FUNCTION_BLOCK TcoContextTest EXTENDS TcoCore._internals_TcoContext
VAR
	_callMyPlcInstance 		:	BOOL := FALSE;
	_startCycles			:	ULINT;
	_endCycles				:	ULINT;	
	_mainCycles				:	ULINT;
	_tcoObjectTest_A		:	TcoObjectTest(THIS^);
	_tcoObjectTest_B		:	TcoObjectTest(THIS^);
	_tcoObjectTest_Misc		:	TcoObjectTest(THIS^);
	_myIdentity				:	ULINT;	
	_onEntryCount			:	ULINT;
	_onExitCount			:	ULINT;
END_VAR

IF THIS^._callMyPlcInstance THEN
	THIS^.Run();
END_IF

{attribute 'TcRpcEnable'}
METHOD INTERNAL CallMainFromUnitTest
THIS^.Main();
END_METHOD

{attribute 'TcRpcEnable'}
METHOD INTERNAL CallRunFromUnitTest
THIS^.Run();
END_METHOD

{attribute 'TcRpcEnable'}
METHOD INTERNAL ContextClose
SUPER^._Close();
END_METHOD

{attribute 'TcRpcEnable'}
METHOD INTERNAL ContextOpen
SUPER^._Open();
END_METHOD

METHOD PROTECTED  Main
_mainCycles := _mainCycles + 1;

_myIdentity	:= THIS^.Identity;
END_METHOD

(*~
	<docu>
		<summary>
			Called on entry into context. When overridden in derived class allows to execute an arbitrary logic prior to opening the context cycle.
			<remarks>			
				<note type="important">					
					The method executes prior to opening the context. The context might not be properly initialized on first call. 
					Any information contained in the context at this point are from the last execution.
				</note>
			</remarks>
		</summary>			
	</docu>	
~*)
METHOD PROTECTED OnEntry
_onEntryCount := _onEntryCount + 1;
END_METHOD


(*~
	<docu>
		<summary>
			Called upon exit from the context. When overridden in derived class allows to execute an arbitrary logic after closing the context cycle.	
		</summary>			
	</docu>	
~*)METHOD PROTECTED OnExit
_onExitCount := _onExitCount + 1;
END_METHOD

{attribute 'TcRpcEnable'}
METHOD INTERNAL ReadOutCycleCounters
_startCycles		:=		THIS^.StartCycleCount;
_endCycles			:=		THIS^.EndCycleCount;

_myIdentity			:= 		THIS^.Identity;
END_METHOD

END_FUNCTION_BLOCK

(* stored: Version 1.1.0.1
   POU TcoContextTest: Id {6642835d-5414-4760-aac1-4c8cef083deb}, SpecialFunc None
   Method CallMainFromUnitTest: Id {9c9d295d-40fb-48af-adaf-5d210f5656a3}
   Method CallRunFromUnitTest: Id {06319017-0b6a-4225-bce8-de1fd8b0ed0e}
   Method ContextClose: Id {4adc0216-d7dc-47d4-a216-4cfc4c14ed41}
   Method ContextOpen: Id {65cd14ad-eb62-4d0c-8ca2-8e3c5c9380bf}
   Method Main: Id {76d8f63c-d45d-4de4-ad73-4298aca95aa1}
   Method OnEntry: Id {39b0dbf1-f025-08a9-2dd6-50f0eee94985}
   Method OnExit: Id {4d6a4e29-82b5-0f04-0eb3-ca65f1c618ae}
   Method ReadOutCycleCounters: Id {3ce97aaa-6bf5-4a06-9e7c-0d88acee2466} *)
